Fanuc KAREL source: KT00534.KL

PROGRAM KT00534
%NOLOCKGROUP
VAR
  P1: JOINTPOS
  P2: POSITION
  OUT: POSITION
BEGIN
  OUT = P1 : P2
END KT00534
